Fanuc KAREL source: kt00244.KL

-- PROVISIONAL review KL for V770-1; original PC SHA256 6a8c9cf9ddaa74489fbb3c71f8bf2924436401fe0166734095b1ccbfa12a6fda
-- Incomplete behavior may be omitted. Consult companion uncertainty JSON. Do not deploy.
PROGRAM KT00244
%NOLOCKGROUP
VAR
  I2 : INTEGER
  OUT : INTEGER
-- UNRESOLVED_DECL Y1 type=002018
BEGIN
  -- UNRESOLVED_PC offsets 5-19; opcodes 2E,22,9D,33,B2
  -- UNRESOLVED_PC offsets 24-35; opcodes 2E,23
  -- UNRESOLVED_PC offsets 40-62; opcodes 22,9D,33,B1,21,47,23
  -- UNRESOLVED_PC offsets 67-71; opcodes 7F
END KT00244
